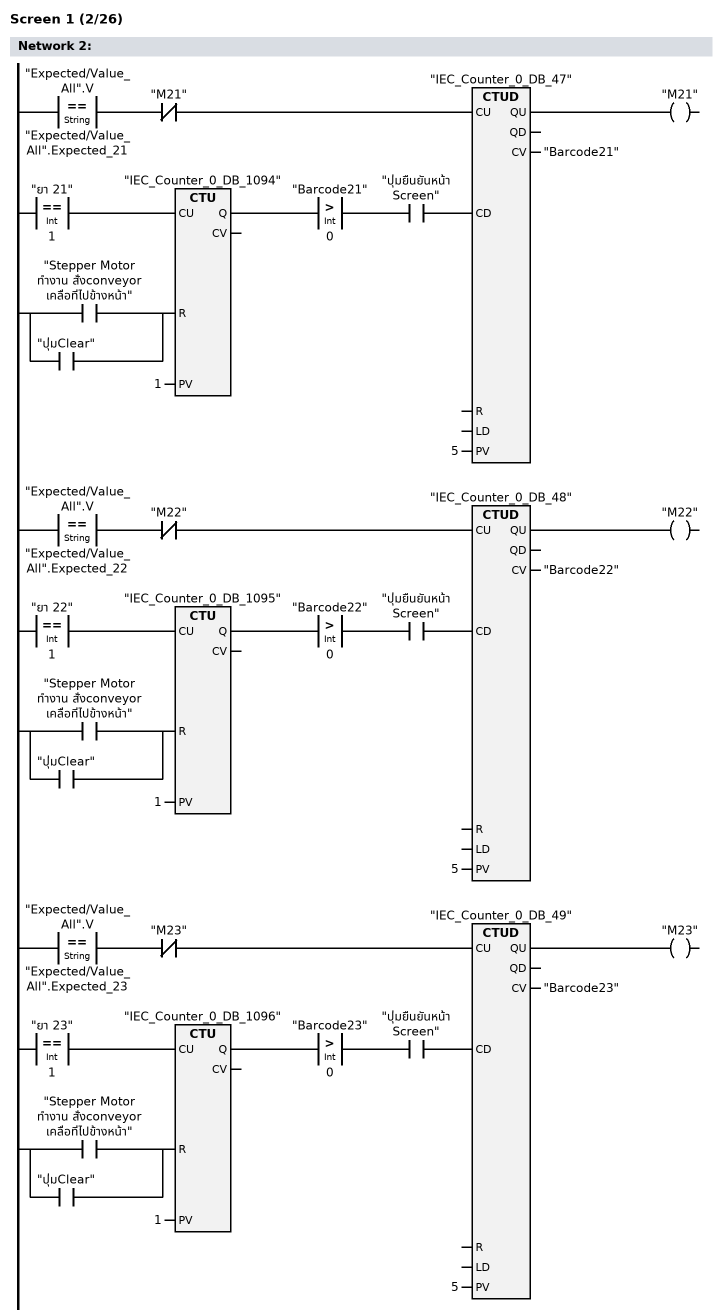
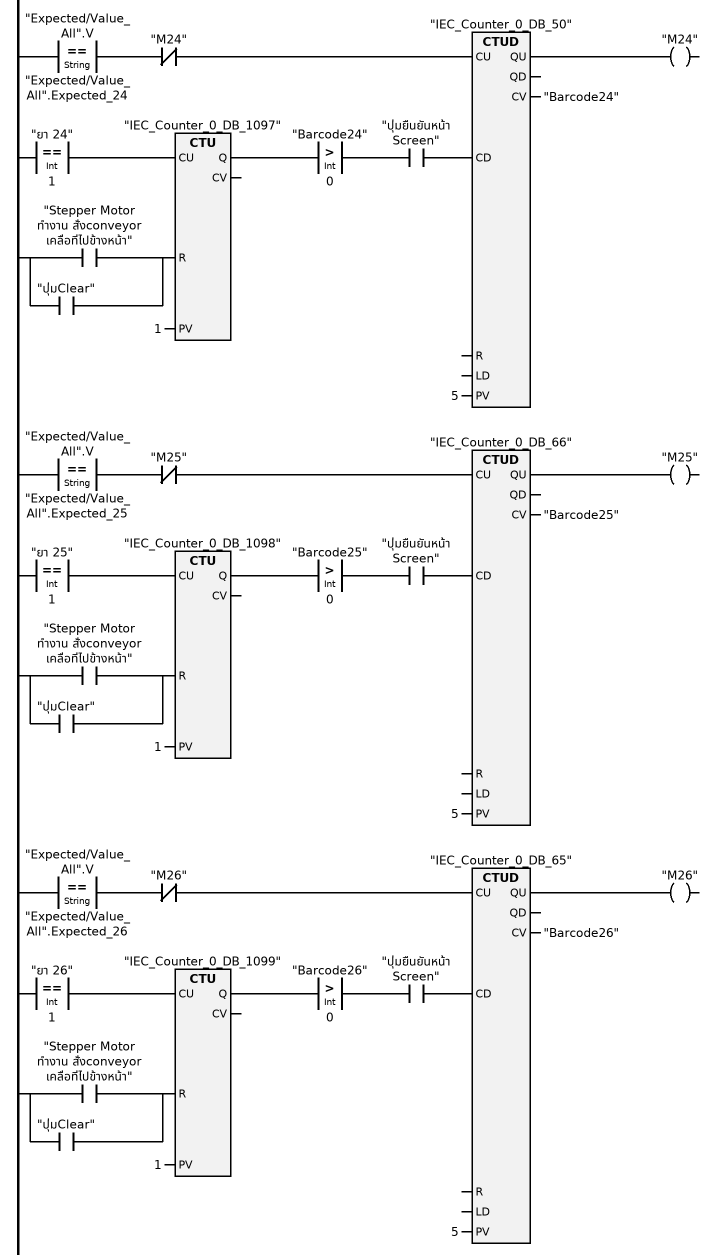
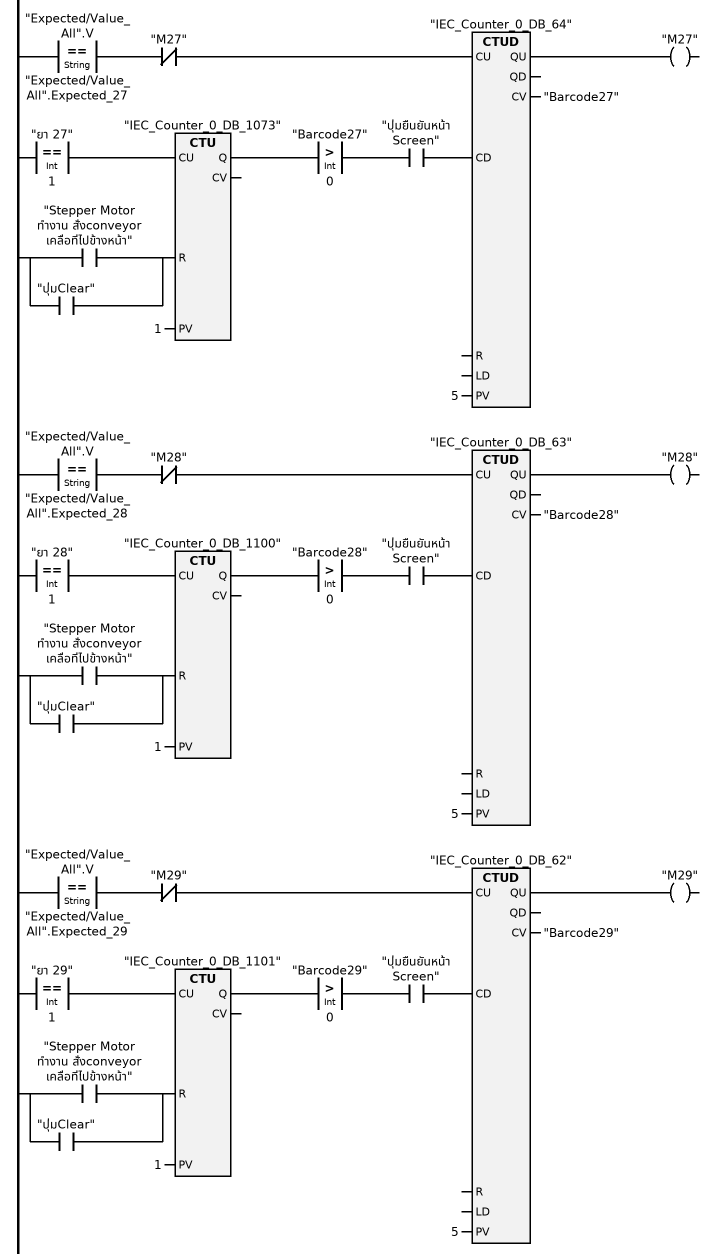
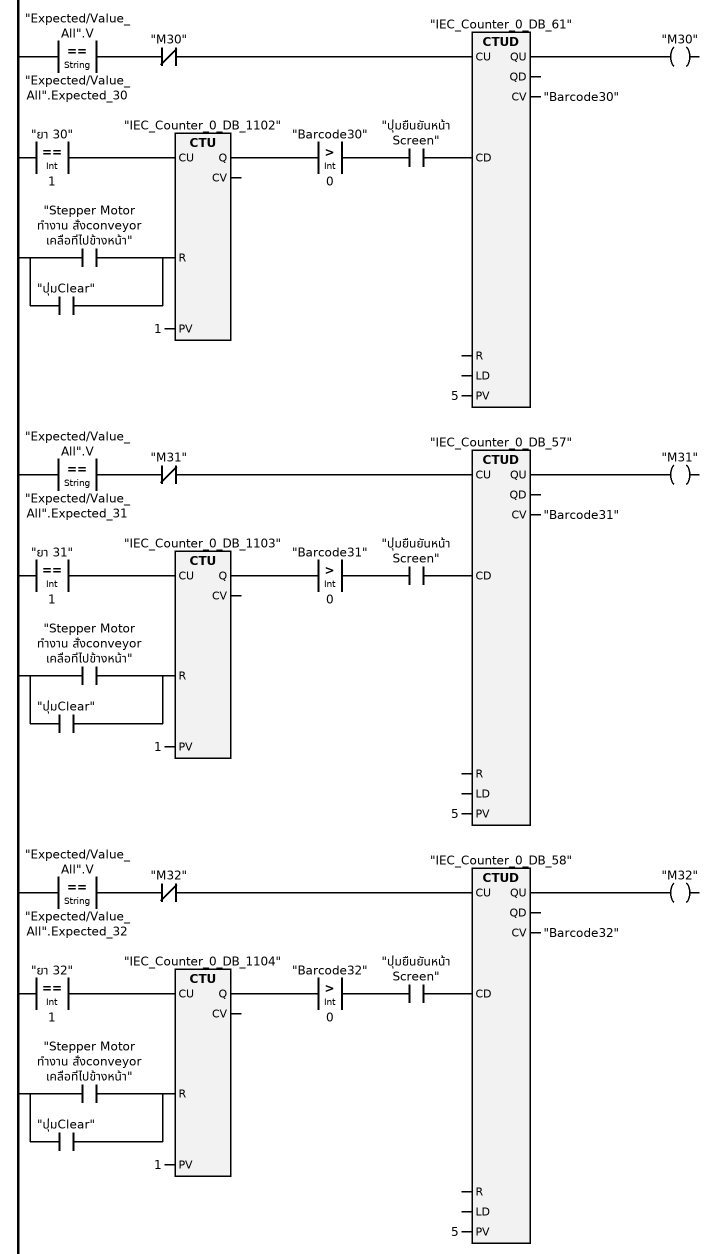
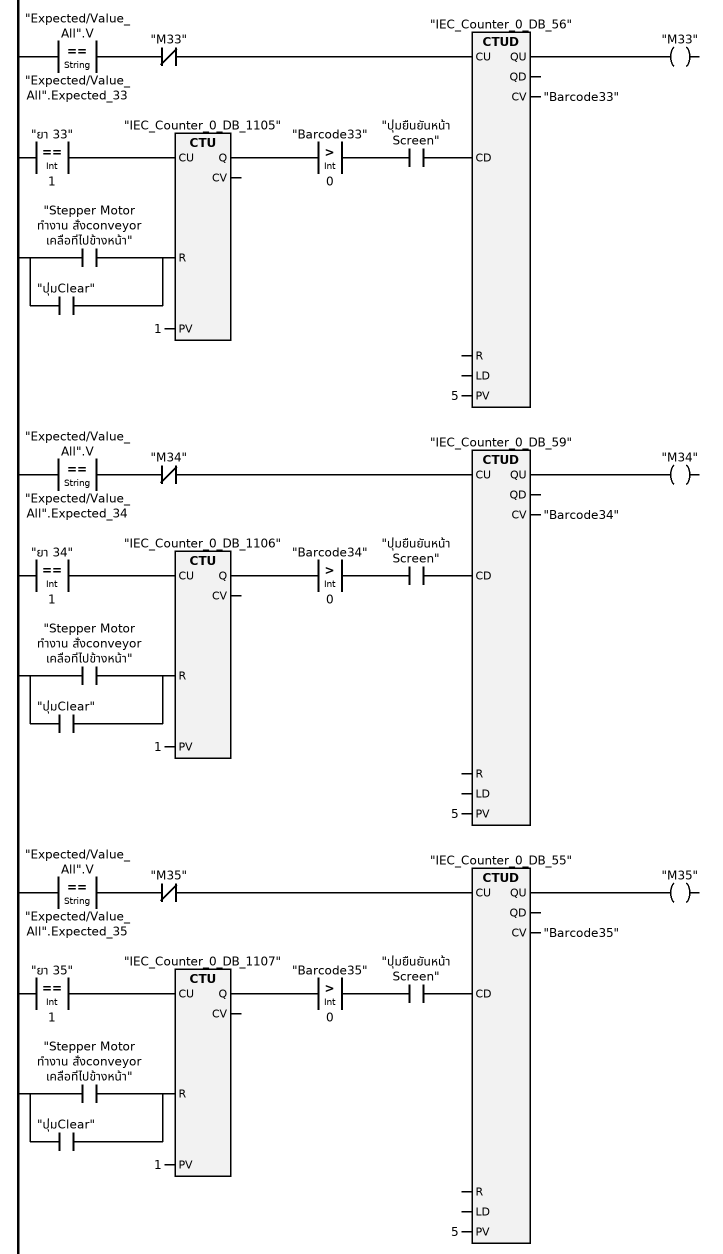
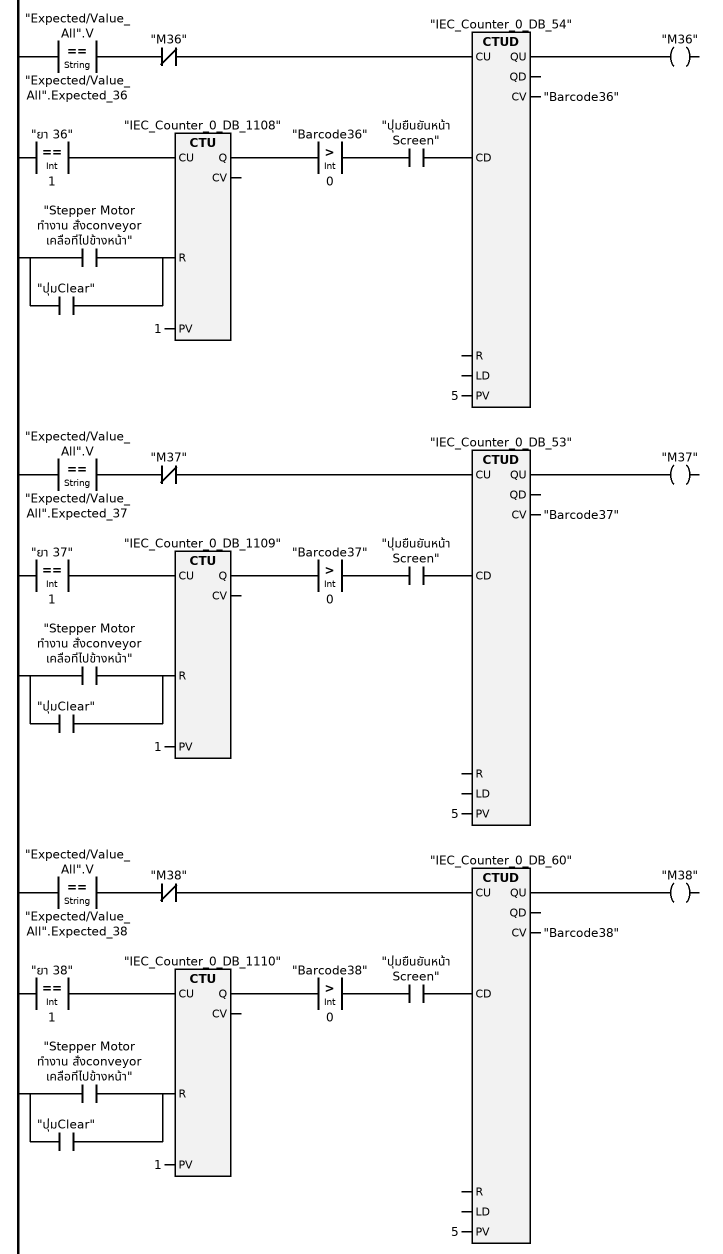
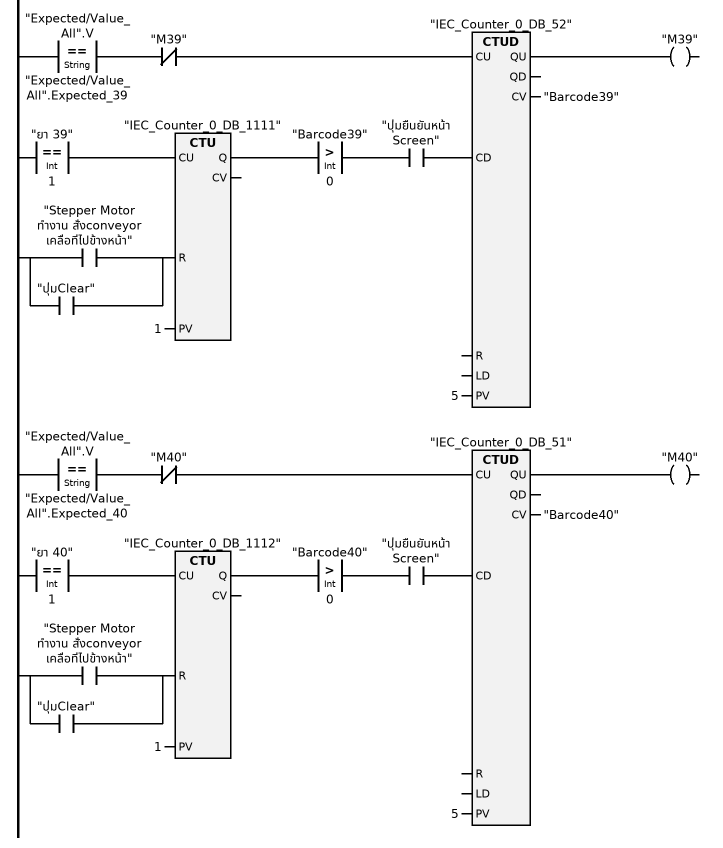
   "IEC_Counter_0_DB_1094".CTU(CU := "ยา 21" = 1,
                           R := "Stepper Motor ทำงาน สั่งconveyor เคลื่อที่ไปข้างหน้า" OR "ปุ่มClear",
                           PV := 1);
   "IEC_Counter_0_DB_47".CTUD(CU := ("Expected/Value_All".V = "Expected/Value_All".Expected_21) AND NOT "M21",
                           CD := "IEC_Counter_0_DB_1094".Q AND ("Barcode21" > 0) AND "ปุ่มยืนยันหน้า Screen",
                           PV := 5,
                           CV => "Barcode21");
   "M21" := "IEC_Counter_0_DB_47".QU;
   "IEC_Counter_0_DB_1095".CTU(CU := "ยา 22" = 1,
                           R := "Stepper Motor ทำงาน สั่งconveyor เคลื่อที่ไปข้างหน้า" OR "ปุ่มClear",
                           PV := 1);
   "IEC_Counter_0_DB_48".CTUD(CU := ("Expected/Value_All".V = "Expected/Value_All".Expected_22) AND NOT "M22",
                           CD := "IEC_Counter_0_DB_1095".Q AND ("Barcode22" > 0) AND "ปุ่มยืนยันหน้า Screen",
                           PV := 5,
                           CV => "Barcode22");
   "M22" := "IEC_Counter_0_DB_48".QU;
   "IEC_Counter_0_DB_1096".CTU(CU := "ยา 23" = 1,
                           R := "Stepper Motor ทำงาน สั่งconveyor เคลื่อที่ไปข้างหน้า" OR "ปุ่มClear",
                           PV := 1);
   "IEC_Counter_0_DB_49".CTUD(CU := ("Expected/Value_All".V = "Expected/Value_All".Expected_23) AND NOT "M23",
                           CD := "IEC_Counter_0_DB_1096".Q AND ("Barcode23" > 0) AND "ปุ่มยืนยันหน้า Screen",
                           PV := 5,
                           CV => "Barcode23");
   "M23" := "IEC_Counter_0_DB_49".QU;
   "IEC_Counter_0_DB_1097".CTU(CU := "ยา 24" = 1,
                           R := "Stepper Motor ทำงาน สั่งconveyor เคลื่อที่ไปข้างหน้า" OR "ปุ่มClear",
                           PV := 1);
   "IEC_Counter_0_DB_50".CTUD(CU := ("Expected/Value_All".V = "Expected/Value_All".Expected_24) AND NOT "M24",
                           CD := "IEC_Counter_0_DB_1097".Q AND ("Barcode24" > 0) AND "ปุ่มยืนยันหน้า Screen",
                           PV := 5,
                           CV => "Barcode24");
   "M24" := "IEC_Counter_0_DB_50".QU;
   "IEC_Counter_0_DB_1098".CTU(CU := "ยา 25" = 1,
                           R := "Stepper Motor ทำงาน สั่งconveyor เคลื่อที่ไปข้างหน้า" OR "ปุ่มClear",
                           PV := 1);
   "IEC_Counter_0_DB_66".CTUD(CU := ("Expected/Value_All".V = "Expected/Value_All".Expected_25) AND NOT "M25",
                           CD := "IEC_Counter_0_DB_1098".Q AND ("Barcode25" > 0) AND "ปุ่มยืนยันหน้า Screen",
                           PV := 5,
                           CV => "Barcode25");
   "M25" := "IEC_Counter_0_DB_66".QU;
   "IEC_Counter_0_DB_1099".CTU(CU := "ยา 26" = 1,
                           R := "Stepper Motor ทำงาน สั่งconveyor เคลื่อที่ไปข้างหน้า" OR "ปุ่มClear",
                           PV := 1);
   "IEC_Counter_0_DB_65".CTUD(CU := ("Expected/Value_All".V = "Expected/Value_All".Expected_26) AND NOT "M26",
                           CD := "IEC_Counter_0_DB_1099".Q AND ("Barcode26" > 0) AND "ปุ่มยืนยันหน้า Screen",
                           PV := 5,
                           CV => "Barcode26");
   "M26" := "IEC_Counter_0_DB_65".QU;
   "IEC_Counter_0_DB_1073".CTU(CU := "ยา 27" = 1,
                           R := "Stepper Motor ทำงาน สั่งconveyor เคลื่อที่ไปข้างหน้า" OR "ปุ่มClear",
                           PV := 1);
   "IEC_Counter_0_DB_64".CTUD(CU := ("Expected/Value_All".V = "Expected/Value_All".Expected_27) AND NOT "M27",
                           CD := "IEC_Counter_0_DB_1073".Q AND ("Barcode27" > 0) AND "ปุ่มยืนยันหน้า Screen",
                           PV := 5,
                           CV => "Barcode27");
   "M27" := "IEC_Counter_0_DB_64".QU;
   "IEC_Counter_0_DB_1100".CTU(CU := "ยา 28" = 1,
                           R := "Stepper Motor ทำงาน สั่งconveyor เคลื่อที่ไปข้างหน้า" OR "ปุ่มClear",
                           PV := 1);
   "IEC_Counter_0_DB_63".CTUD(CU := ("Expected/Value_All".V = "Expected/Value_All".Expected_28) AND NOT "M28",
                           CD := "IEC_Counter_0_DB_1100".Q AND ("Barcode28" > 0) AND "ปุ่มยืนยันหน้า Screen",
                           PV := 5,
                           CV => "Barcode28");
   "M28" := "IEC_Counter_0_DB_63".QU;
   "IEC_Counter_0_DB_1101".CTU(CU := "ยา 29" = 1,
                           R := "Stepper Motor ทำงาน สั่งconveyor เคลื่อที่ไปข้างหน้า" OR "ปุ่มClear",
                           PV := 1);
   "IEC_Counter_0_DB_62".CTUD(CU := ("Expected/Value_All".V = "Expected/Value_All".Expected_29) AND NOT "M29",
                           CD := "IEC_Counter_0_DB_1101".Q AND ("Barcode29" > 0) AND "ปุ่มยืนยันหน้า Screen",
                           PV := 5,
                           CV => "Barcode29");
   "M29" := "IEC_Counter_0_DB_62".QU;
   "IEC_Counter_0_DB_1102".CTU(CU := "ยา 30" = 1,
                           R := "Stepper Motor ทำงาน สั่งconveyor เคลื่อที่ไปข้างหน้า" OR "ปุ่มClear",
                           PV := 1);
   "IEC_Counter_0_DB_61".CTUD(CU := ("Expected/Value_All".V = "Expected/Value_All".Expected_30) AND NOT "M30",
                           CD := "IEC_Counter_0_DB_1102".Q AND ("Barcode30" > 0) AND "ปุ่มยืนยันหน้า Screen",
                           PV := 5,
                           CV => "Barcode30");
   "M30" := "IEC_Counter_0_DB_61".QU;
   "IEC_Counter_0_DB_1103".CTU(CU := "ยา 31" = 1,
                           R := "Stepper Motor ทำงาน สั่งconveyor เคลื่อที่ไปข้างหน้า" OR "ปุ่มClear",
                           PV := 1);
   "IEC_Counter_0_DB_57".CTUD(CU := ("Expected/Value_All".V = "Expected/Value_All".Expected_31) AND NOT "M31",
                           CD := "IEC_Counter_0_DB_1103".Q AND ("Barcode31" > 0) AND "ปุ่มยืนยันหน้า Screen",
                           PV := 5,
                           CV => "Barcode31");
   "M31" := "IEC_Counter_0_DB_57".QU;
   "IEC_Counter_0_DB_1104".CTU(CU := "ยา 32" = 1,
                           R := "Stepper Motor ทำงาน สั่งconveyor เคลื่อที่ไปข้างหน้า" OR "ปุ่มClear",
                           PV := 1);
   "IEC_Counter_0_DB_58".CTUD(CU := ("Expected/Value_All".V = "Expected/Value_All".Expected_32) AND NOT "M32",
                           CD := "IEC_Counter_0_DB_1104".Q AND ("Barcode32" > 0) AND "ปุ่มยืนยันหน้า Screen",
                           PV := 5,
                           CV => "Barcode32");
   "M32" := "IEC_Counter_0_DB_58".QU;
   "IEC_Counter_0_DB_1105".CTU(CU := "ยา 33" = 1,
                           R := "Stepper Motor ทำงาน สั่งconveyor เคลื่อที่ไปข้างหน้า" OR "ปุ่มClear",
                           PV := 1);
   "IEC_Counter_0_DB_56".CTUD(CU := ("Expected/Value_All".V = "Expected/Value_All".Expected_33) AND NOT "M33",
                           CD := "IEC_Counter_0_DB_1105".Q AND ("Barcode33" > 0) AND "ปุ่มยืนยันหน้า Screen",
                           PV := 5,
                           CV => "Barcode33");
   "M33" := "IEC_Counter_0_DB_56".QU;
   "IEC_Counter_0_DB_1106".CTU(CU := "ยา 34" = 1,
                           R := "Stepper Motor ทำงาน สั่งconveyor เคลื่อที่ไปข้างหน้า" OR "ปุ่มClear",
                           PV := 1);
   "IEC_Counter_0_DB_59".CTUD(CU := ("Expected/Value_All".V = "Expected/Value_All".Expected_34) AND NOT "M34",
                           CD := "IEC_Counter_0_DB_1106".Q AND ("Barcode34" > 0) AND "ปุ่มยืนยันหน้า Screen",
                           PV := 5,
                           CV => "Barcode34");
   "M34" := "IEC_Counter_0_DB_59".QU;
   "IEC_Counter_0_DB_1107".CTU(CU := "ยา 35" = 1,
                           R := "Stepper Motor ทำงาน สั่งconveyor เคลื่อที่ไปข้างหน้า" OR "ปุ่มClear",
                           PV := 1);
   "IEC_Counter_0_DB_55".CTUD(CU := ("Expected/Value_All".V = "Expected/Value_All".Expected_35) AND NOT "M35",
                           CD := "IEC_Counter_0_DB_1107".Q AND ("Barcode35" > 0) AND "ปุ่มยืนยันหน้า Screen",
                           PV := 5,
                           CV => "Barcode35");
   "M35" := "IEC_Counter_0_DB_55".QU;
   "IEC_Counter_0_DB_1108".CTU(CU := "ยา 36" = 1,
                           R := "Stepper Motor ทำงาน สั่งconveyor เคลื่อที่ไปข้างหน้า" OR "ปุ่มClear",
                           PV := 1);
   "IEC_Counter_0_DB_54".CTUD(CU := ("Expected/Value_All".V = "Expected/Value_All".Expected_36) AND NOT "M36",
                           CD := "IEC_Counter_0_DB_1108".Q AND ("Barcode36" > 0) AND "ปุ่มยืนยันหน้า Screen",
                           PV := 5,
                           CV => "Barcode36");
   "M36" := "IEC_Counter_0_DB_54".QU;
   "IEC_Counter_0_DB_1109".CTU(CU := "ยา 37" = 1,
                           R := "Stepper Motor ทำงาน สั่งconveyor เคลื่อที่ไปข้างหน้า" OR "ปุ่มClear",
                           PV := 1);
   "IEC_Counter_0_DB_53".CTUD(CU := ("Expected/Value_All".V = "Expected/Value_All".Expected_37) AND NOT "M37",
                           CD := "IEC_Counter_0_DB_1109".Q AND ("Barcode37" > 0) AND "ปุ่มยืนยันหน้า Screen",
                           PV := 5,
                           CV => "Barcode37");
   "M37" := "IEC_Counter_0_DB_53".QU;
   "IEC_Counter_0_DB_1110".CTU(CU := "ยา 38" = 1,
                           R := "Stepper Motor ทำงาน สั่งconveyor เคลื่อที่ไปข้างหน้า" OR "ปุ่มClear",
                           PV := 1);
   "IEC_Counter_0_DB_60".CTUD(CU := ("Expected/Value_All".V = "Expected/Value_All".Expected_38) AND NOT "M38",
                           CD := "IEC_Counter_0_DB_1110".Q AND ("Barcode38" > 0) AND "ปุ่มยืนยันหน้า Screen",
                           PV := 5,
                           CV => "Barcode38");
   "M38" := "IEC_Counter_0_DB_60".QU;
   "IEC_Counter_0_DB_1111".CTU(CU := "ยา 39" = 1,
                           R := "Stepper Motor ทำงาน สั่งconveyor เคลื่อที่ไปข้างหน้า" OR "ปุ่มClear",
                           PV := 1);
   "IEC_Counter_0_DB_52".CTUD(CU := ("Expected/Value_All".V = "Expected/Value_All".Expected_39) AND NOT "M39",
                           CD := "IEC_Counter_0_DB_1111".Q AND ("Barcode39" > 0) AND "ปุ่มยืนยันหน้า Screen",
                           PV := 5,
                           CV => "Barcode39");
   "M39" := "IEC_Counter_0_DB_52".QU;
   "IEC_Counter_0_DB_1112".CTU(CU := "ยา 40" = 1,
                           R := "Stepper Motor ทำงาน สั่งconveyor เคลื่อที่ไปข้างหน้า" OR "ปุ่มClear",
                           PV := 1);
   "IEC_Counter_0_DB_51".CTUD(CU := ("Expected/Value_All".V = "Expected/Value_All".Expected_40) AND NOT "M40",
                           CD := "IEC_Counter_0_DB_1112".Q AND ("Barcode40" > 0) AND "ปุ่มยืนยันหน้า Screen",
                           PV := 5,
                           CV => "Barcode40");
   "M40" := "IEC_Counter_0_DB_51".QU;
END_REGION

REGION Network 3
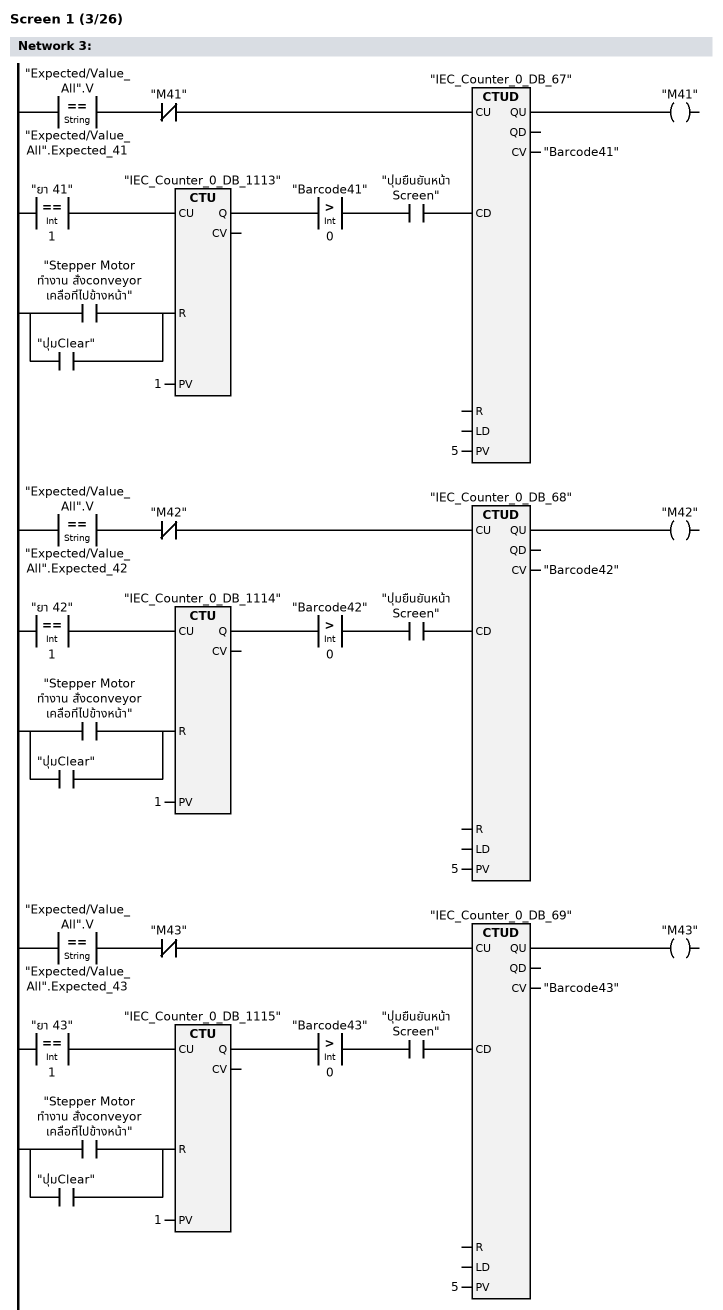
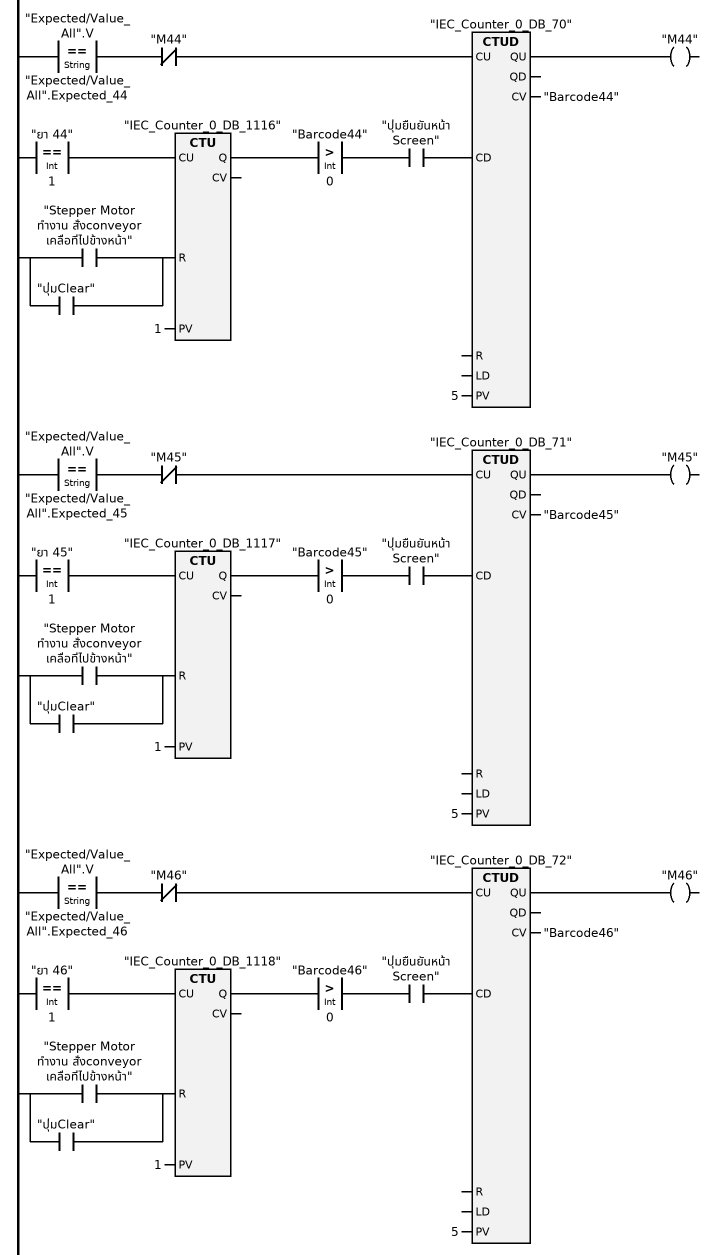
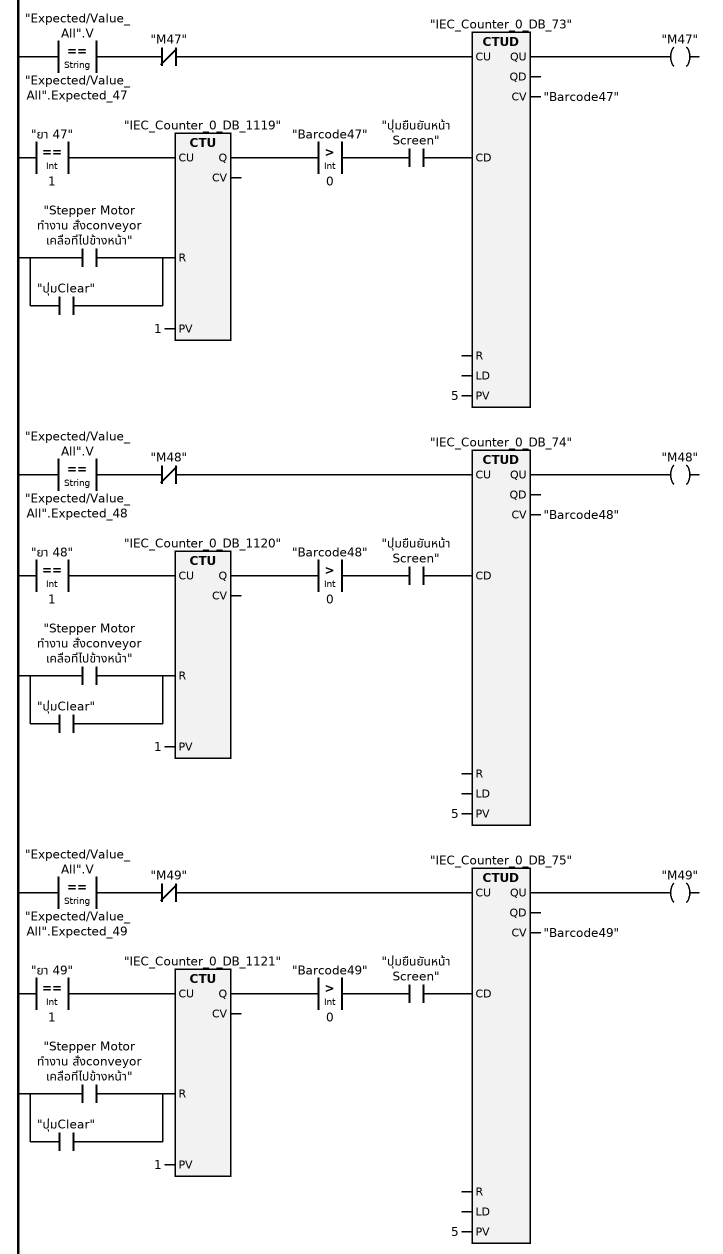
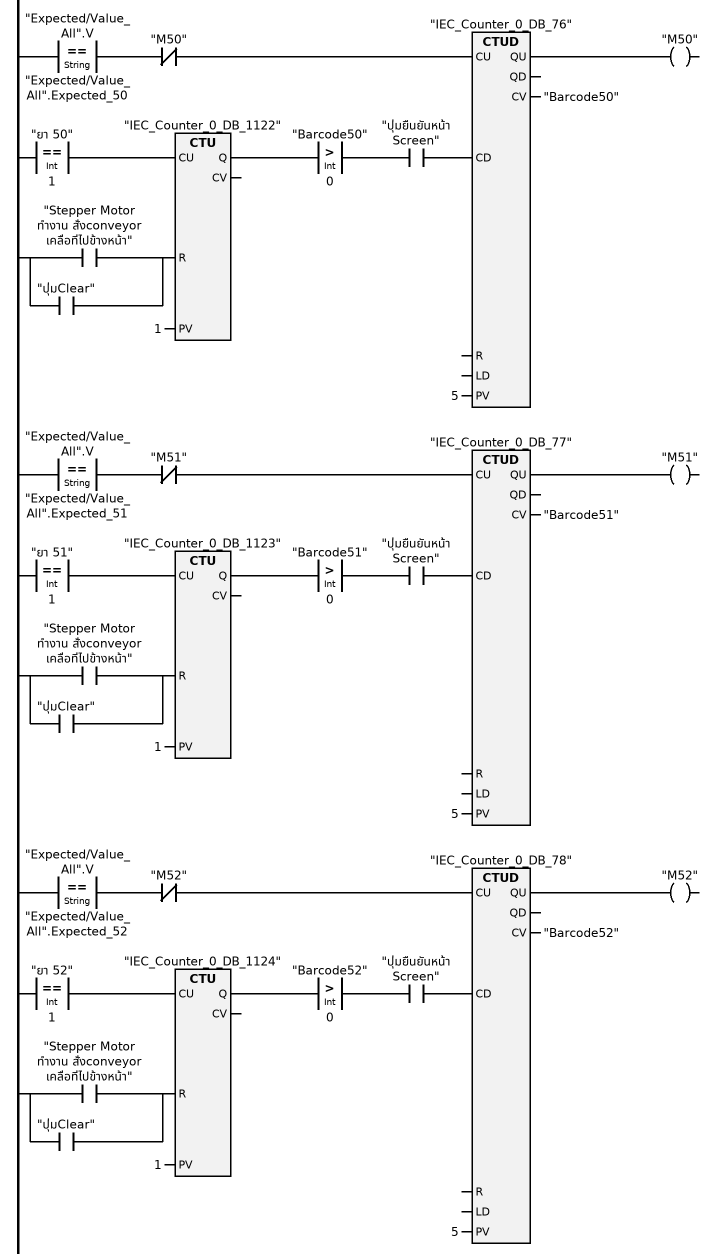
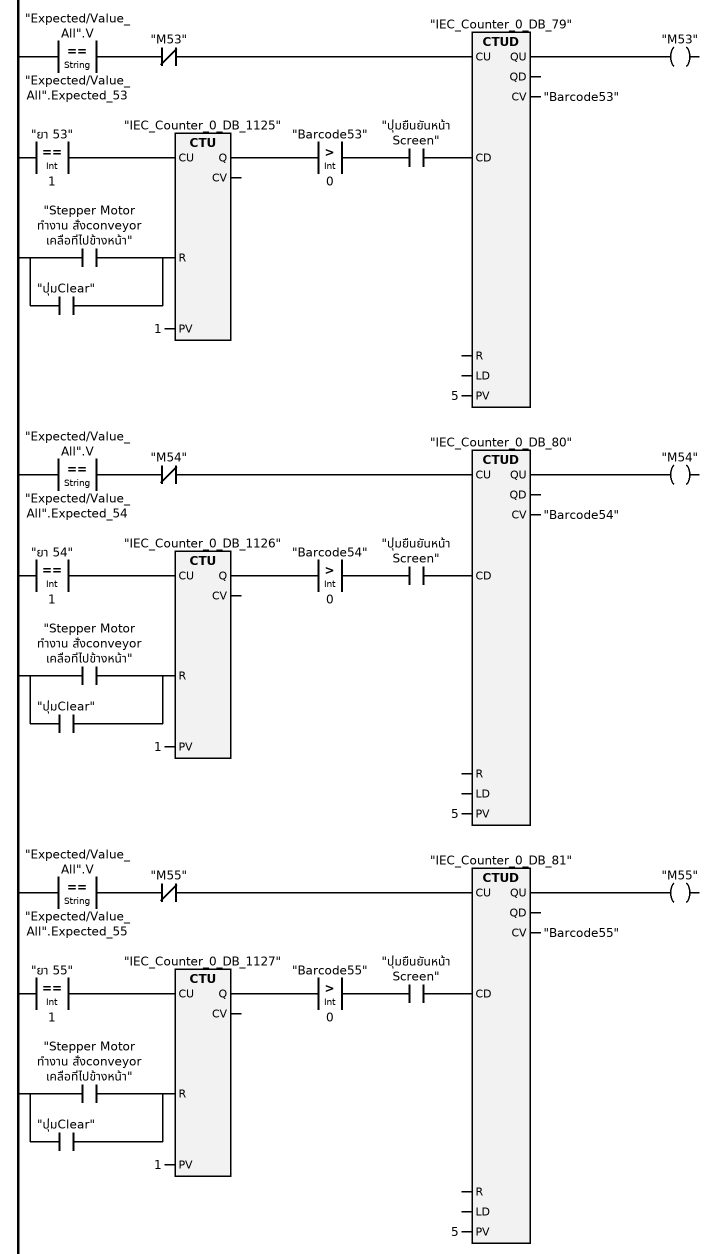
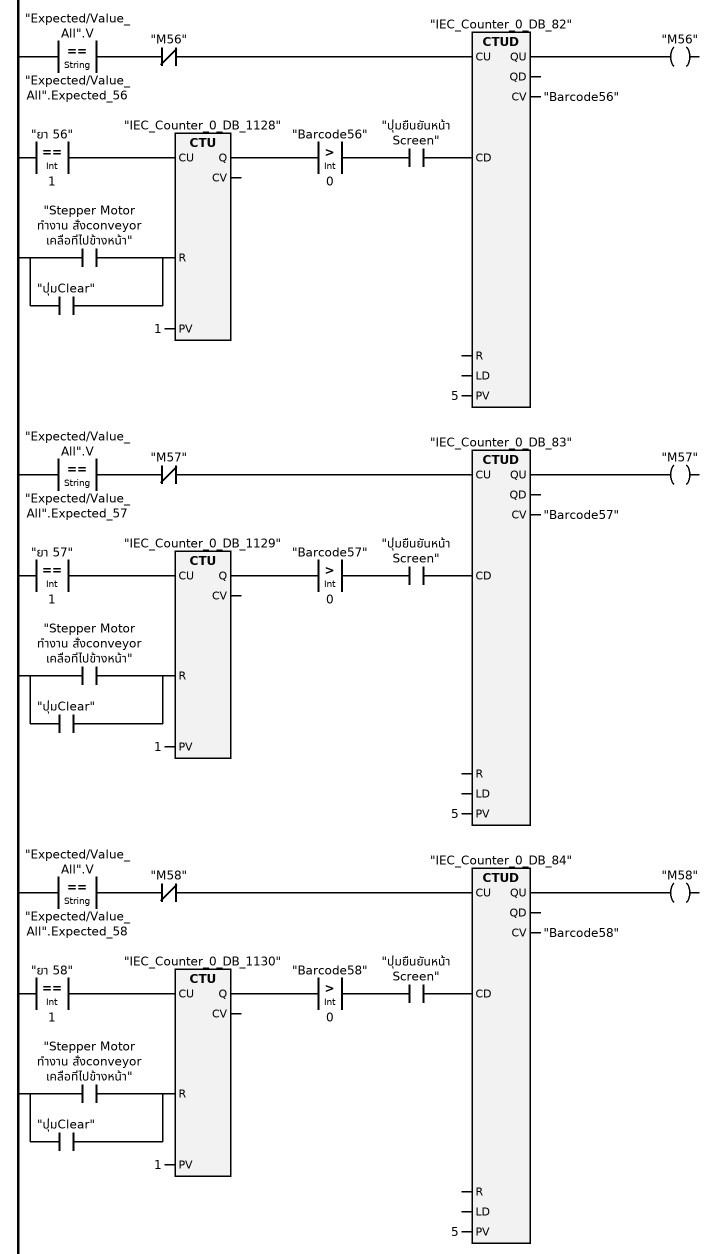
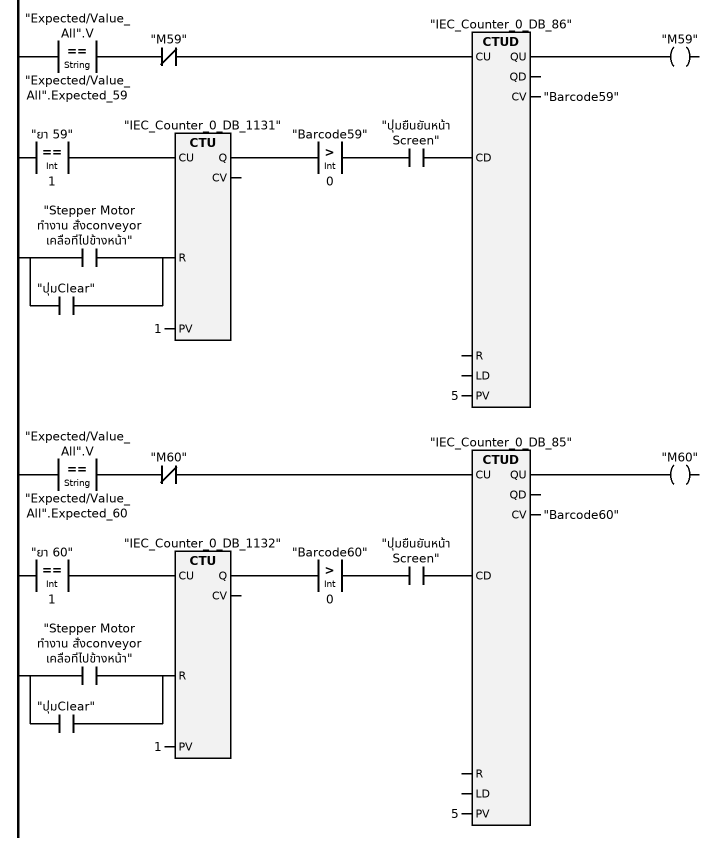
   "IEC_Counter_0_DB_1113".CTU(CU := "ยา 41" = 1,
                           R := "Stepper Motor ทำงาน สั่งconveyor เคลื่อที่ไปข้างหน้า" OR "ปุ่มClear",
                           PV := 1);
   "IEC_Counter_0_DB_67".CTUD(CU := ("Expected/Value_All".V = "Expected/Value_All".Expected_41) AND NOT "M41",
                           CD := "IEC_Counter_0_DB_1113".Q AND ("Barcode41" > 0) AND "ปุ่มยืนยันหน้า Screen",
                           PV := 5,
                           CV => "Barcode41");
   "M41" := "IEC_Counter_0_DB_67".QU;
   "IEC_Counter_0_DB_1114".CTU(CU := "ยา 42" = 1,
                           R := "Stepper Motor ทำงาน สั่งconveyor เคลื่อที่ไปข้างหน้า" OR "ปุ่มClear",
                           PV := 1);
   "IEC_Counter_0_DB_68".CTUD(CU := ("Expected/Value_All".V = "Expected/Value_All".Expected_42) AND NOT "M42",
                           CD := "IEC_Counter_0_DB_1114".Q AND ("Barcode42" > 0) AND "ปุ่มยืนยันหน้า Screen",
                           PV := 5,
                           CV => "Barcode42");
   "M42" := "IEC_Counter_0_DB_68".QU;
   "IEC_Counter_0_DB_1115".CTU(CU := "ยา 43" = 1,
                           R := "Stepper Motor ทำงาน สั่งconveyor เคลื่อที่ไปข้างหน้า" OR "ปุ่มClear",
                           PV := 1);
   "IEC_Counter_0_DB_69".CTUD(CU := ("Expected/Value_All".V = "Expected/Value_All".Expected_43) AND NOT "M43",
                           CD := "IEC_Counter_0_DB_1115".Q AND ("Barcode43" > 0) AND "ปุ่มยืนยันหน้า Screen",
                           PV := 5,
                           CV => "Barcode43");
   "M43" := "IEC_Counter_0_DB_69".QU;
   "IEC_Counter_0_DB_1116".CTU(CU := "ยา 44" = 1,
                           R := "Stepper Motor ทำงาน สั่งconveyor เคลื่อที่ไปข้างหน้า" OR "ปุ่มClear",
                           PV := 1);
   "IEC_Counter_0_DB_70".CTUD(CU := ("Expected/Value_All".V = "Expected/Value_All".Expected_44) AND NOT "M44",
                           CD := "IEC_Counter_0_DB_1116".Q AND ("Barcode44" > 0) AND "ปุ่มยืนยันหน้า Screen",
                           PV := 5,
                           CV => "Barcode44");
   "M44" := "IEC_Counter_0_DB_70".QU;
   "IEC_Counter_0_DB_1117".CTU(CU := "ยา 45" = 1,
                           R := "Stepper Motor ทำงาน สั่งconveyor เคลื่อที่ไปข้างหน้า" OR "ปุ่มClear",
                           PV := 1);
   "IEC_Counter_0_DB_71".CTUD(CU := ("Expected/Value_All".V = "Expected/Value_All".Expected_45) AND NOT "M45",
                           CD := "IEC_Counter_0_DB_1117".Q AND ("Barcode45" > 0) AND "ปุ่มยืนยันหน้า Screen",
                           PV := 5,
                           CV => "Barcode45");
   "M45" := "IEC_Counter_0_DB_71".QU;
   "IEC_Counter_0_DB_1118".CTU(CU := "ยา 46" = 1,
                           R := "Stepper Motor ทำงาน สั่งconveyor เคลื่อที่ไปข้างหน้า" OR "ปุ่มClear",
                           PV := 1);
   "IEC_Counter_0_DB_72".CTUD(CU := ("Expected/Value_All".V = "Expected/Value_All".Expected_46) AND NOT "M46",
                           CD := "IEC_Counter_0_DB_1118".Q AND ("Barcode46" > 0) AND "ปุ่มยืนยันหน้า Screen",
                           PV := 5,
                           CV => "Barcode46");
   "M46" := "IEC_Counter_0_DB_72".QU;
   "IEC_Counter_0_DB_1119".CTU(CU := "ยา 47" = 1,
                           R := "Stepper Motor ทำงาน สั่งconveyor เคลื่อที่ไปข้างหน้า" OR "ปุ่มClear",
                           PV := 1);
   "IEC_Counter_0_DB_73".CTUD(CU := ("Expected/Value_All".V = "Expected/Value_All".Expected_47) AND NOT "M47",
                           CD := "IEC_Counter_0_DB_1119".Q AND ("Barcode47" > 0) AND "ปุ่มยืนยันหน้า Screen",
                           PV := 5,
                           CV => "Barcode47");
   "M47" := "IEC_Counter_0_DB_73".QU;
   "IEC_Counter_0_DB_1120".CTU(CU := "ยา 48" = 1,
                           R := "Stepper Motor ทำงาน สั่งconveyor เคลื่อที่ไปข้างหน้า" OR "ปุ่มClear",
                           PV := 1);
   "IEC_Counter_0_DB_74".CTUD(CU := ("Expected/Value_All".V = "Expected/Value_All".Expected_48) AND NOT "M48",
                           CD := "IEC_Counter_0_DB_1120".Q AND ("Barcode48" > 0) AND "ปุ่มยืนยันหน้า Screen",
                           PV := 5,
                           CV => "Barcode48");
   "M48" := "IEC_Counter_0_DB_74".QU;
   "IEC_Counter_0_DB_1121".CTU(CU := "ยา 49" = 1,
                           R := "Stepper Motor ทำงาน สั่งconveyor เคลื่อที่ไปข้างหน้า" OR "ปุ่มClear",
                           PV := 1);
   "IEC_Counter_0_DB_75".CTUD(CU := ("Expected/Value_All".V = "Expected/Value_All".Expected_49) AND NOT "M49",
                           CD := "IEC_Counter_0_DB_1121".Q AND ("Barcode49" > 0) AND "ปุ่มยืนยันหน้า Screen",
                           PV := 5,
                           CV => "Barcode49");
   "M49" := "IEC_Counter_0_DB_75".QU;
   "IEC_Counter_0_DB_1122".CTU(CU := "ยา 50" = 1,
                           R := "Stepper Motor ทำงาน สั่งconveyor เคลื่อที่ไปข้างหน้า" OR "ปุ่มClear",
                           PV := 1);
   "IEC_Counter_0_DB_76".CTUD(CU := ("Expected/Value_All".V = "Expected/Value_All".Expected_50) AND NOT "M50",
                           CD := "IEC_Counter_0_DB_1122".Q AND ("Barcode50" > 0) AND "ปุ่มยืนยันหน้า Screen",
                           PV := 5,
                           CV => "Barcode50");
   "M50" := "IEC_Counter_0_DB_76".QU;
   "IEC_Counter_0_DB_1123".CTU(CU := "ยา 51" = 1,
                           R := "Stepper Motor ทำงาน สั่งconveyor เคลื่อที่ไปข้างหน้า" OR "ปุ่มClear",
                           PV := 1);
   "IEC_Counter_0_DB_77".CTUD(CU := ("Expected/Value_All".V = "Expected/Value_All".Expected_51) AND NOT "M51",
                           CD := "IEC_Counter_0_DB_1123".Q AND ("Barcode51" > 0) AND "ปุ่มยืนยันหน้า Screen",
                           PV := 5,
                           CV => "Barcode51");
   "M51" := "IEC_Counter_0_DB_77".QU;
   "IEC_Counter_0_DB_1124".CTU(CU := "ยา 52" = 1,
                           R := "Stepper Motor ทำงาน สั่งconveyor เคลื่อที่ไปข้างหน้า" OR "ปุ่มClear",
                           PV := 1);
   "IEC_Counter_0_DB_78".CTUD(CU := ("Expected/Value_All".V = "Expected/Value_All".Expected_52) AND NOT "M52",
                           CD := "IEC_Counter_0_DB_1124".Q AND ("Barcode52" > 0) AND "ปุ่มยืนยันหน้า Screen",
                           PV := 5,
                           CV => "Barcode52");
   "M52" := "IEC_Counter_0_DB_78".QU;
   "IEC_Counter_0_DB_1125".CTU(CU := "ยา 53" = 1,
                           R := "Stepper Motor ทำงาน สั่งconveyor เคลื่อที่ไปข้างหน้า" OR "ปุ่มClear",
                           PV := 1);
   "IEC_Counter_0_DB_79".CTUD(CU := ("Expected/Value_All".V = "Expected/Value_All".Expected_53) AND NOT "M53",
                           CD := "IEC_Counter_0_DB_1125".Q AND ("Barcode53" > 0) AND "ปุ่มยืนยันหน้า Screen",
                           PV := 5,
                           CV => "Barcode53");
   "M53" := "IEC_Counter_0_DB_79".QU;
   "IEC_Counter_0_DB_1126".CTU(CU := "ยา 54" = 1,
                           R := "Stepper Motor ทำงาน สั่งconveyor เคลื่อที่ไปข้างหน้า" OR "ปุ่มClear",
                           PV := 1);
   "IEC_Counter_0_DB_80".CTUD(CU := ("Expected/Value_All".V = "Expected/Value_All".Expected_54) AND NOT "M54",
                           CD := "IEC_Counter_0_DB_1126".Q AND ("Barcode54" > 0) AND "ปุ่มยืนยันหน้า Screen",
                           PV := 5,
                           CV => "Barcode54");
   "M54" := "IEC_Counter_0_DB_80".QU;
   "IEC_Counter_0_DB_1127".CTU(CU := "ยา 55" = 1,
                           R := "Stepper Motor ทำงาน สั่งconveyor เคลื่อที่ไปข้างหน้า" OR "ปุ่มClear",
                           PV := 1);
   "IEC_Counter_0_DB_81".CTUD(CU := ("Expected/Value_All".V = "Expected/Value_All".Expected_55) AND NOT "M55",
                           CD := "IEC_Counter_0_DB_1127".Q AND ("Barcode55" > 0) AND "ปุ่มยืนยันหน้า Screen",
                           PV := 5,
                           CV => "Barcode55");
   "M55" := "IEC_Counter_0_DB_81".QU;
   "IEC_Counter_0_DB_1128".CTU(CU := "ยา 56" = 1,
                           R := "Stepper Motor ทำงาน สั่งconveyor เคลื่อที่ไปข้างหน้า" OR "ปุ่มClear",
                           PV := 1);
   "IEC_Counter_0_DB_82".CTUD(CU := ("Expected/Value_All".V = "Expected/Value_All".Expected_56) AND NOT "M56",
                           CD := "IEC_Counter_0_DB_1128".Q AND ("Barcode56" > 0) AND "ปุ่มยืนยันหน้า Screen",
                           PV := 5,
                           CV => "Barcode56");
   "M56" := "IEC_Counter_0_DB_82".QU;
   "IEC_Counter_0_DB_1129".CTU(CU := "ยา 57" = 1,
                           R := "Stepper Motor ทำงาน สั่งconveyor เคลื่อที่ไปข้างหน้า" OR "ปุ่มClear",
                           PV := 1);
   "IEC_Counter_0_DB_83".CTUD(CU := ("Expected/Value_All".V = "Expected/Value_All".Expected_57) AND NOT "M57",
                           CD := "IEC_Counter_0_DB_1129".Q AND ("Barcode57" > 0) AND "ปุ่มยืนยันหน้า Screen",
                           PV := 5,
                           CV => "Barcode57");
   "M57" := "IEC_Counter_0_DB_83".QU;
   "IEC_Counter_0_DB_1130".CTU(CU := "ยา 58" = 1,
                           R := "Stepper Motor ทำงาน สั่งconveyor เคลื่อที่ไปข้างหน้า" OR "ปุ่มClear",
                           PV := 1);
   "IEC_Counter_0_DB_84".CTUD(CU := ("Expected/Value_All".V = "Expected/Value_All".Expected_58) AND NOT "M58",
                           CD := "IEC_Counter_0_DB_1130".Q AND ("Barcode58" > 0) AND "ปุ่มยืนยันหน้า Screen",
                           PV := 5,
                           CV => "Barcode58");
   "M58" := "IEC_Counter_0_DB_84".QU;
   "IEC_Counter_0_DB_1131".CTU(CU := "ยา 59" = 1,
                           R := "Stepper Motor ทำงาน สั่งconveyor เคลื่อที่ไปข้างหน้า" OR "ปุ่มClear",
                           PV := 1);
   "IEC_Counter_0_DB_86".CTUD(CU := ("Expected/Value_All".V = "Expected/Value_All".Expected_59) AND NOT "M59",
                           CD := "IEC_Counter_0_DB_1131".Q AND ("Barcode59" > 0) AND "ปุ่มยืนยันหน้า Screen",
                           PV := 5,
                           CV => "Barcode59");
   "M59" := "IEC_Counter_0_DB_86".QU;
   "IEC_Counter_0_DB_1132".CTU(CU := "ยา 60" = 1,
                           R := "Stepper Motor ทำงาน สั่งconveyor เคลื่อที่ไปข้างหน้า" OR "ปุ่มClear",
                           PV := 1);
   "IEC_Counter_0_DB_85".CTUD(CU := ("Expected/Value_All".V = "Expected/Value_All".Expected_60) AND NOT "M60",
                           CD := "IEC_Counter_0_DB_1132".Q AND ("Barcode60" > 0) AND "ปุ่มยืนยันหน้า Screen",
                           PV := 5,
                           CV => "Barcode60");
   "M60" := "IEC_Counter_0_DB_85".QU;
END_REGION

REGION Network 4
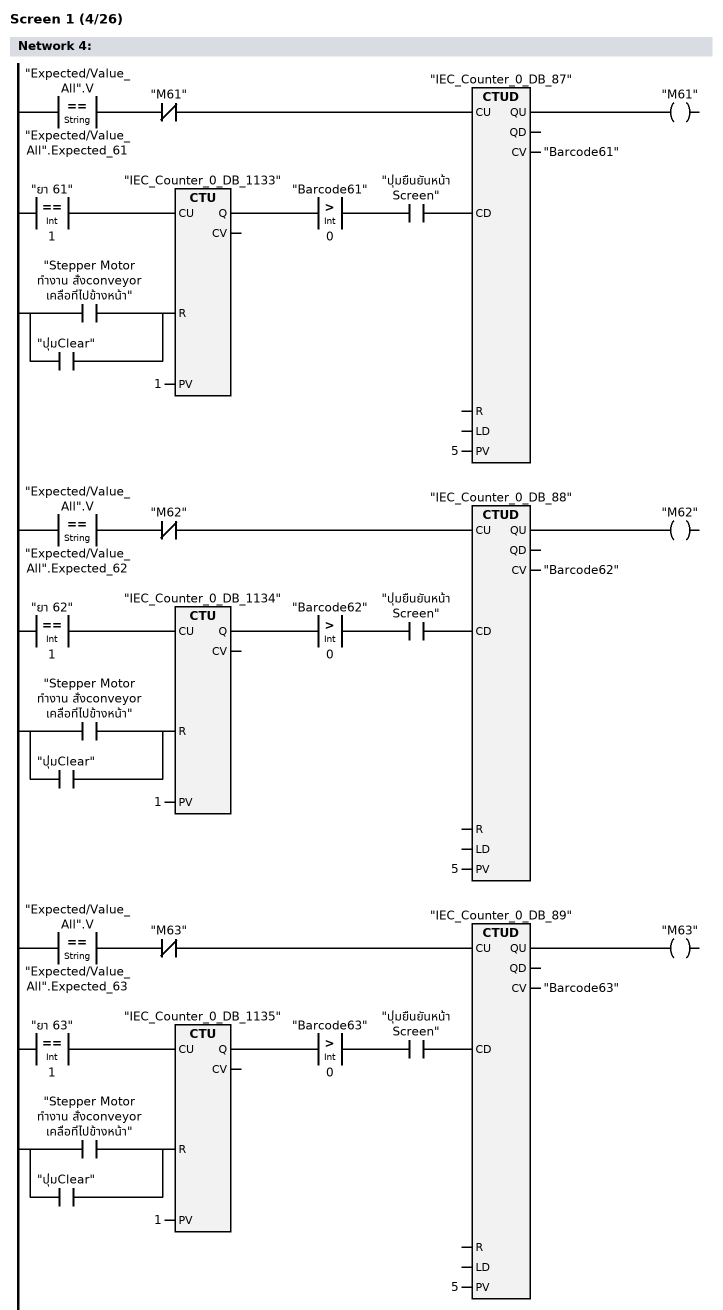
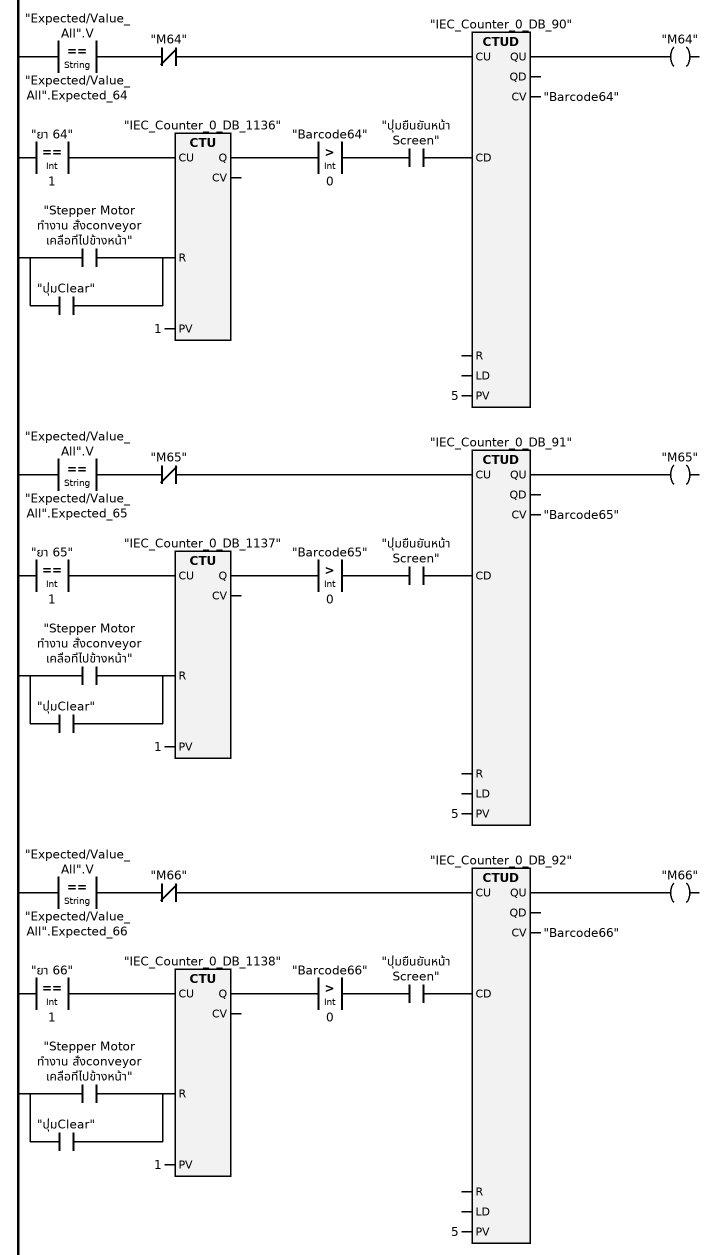
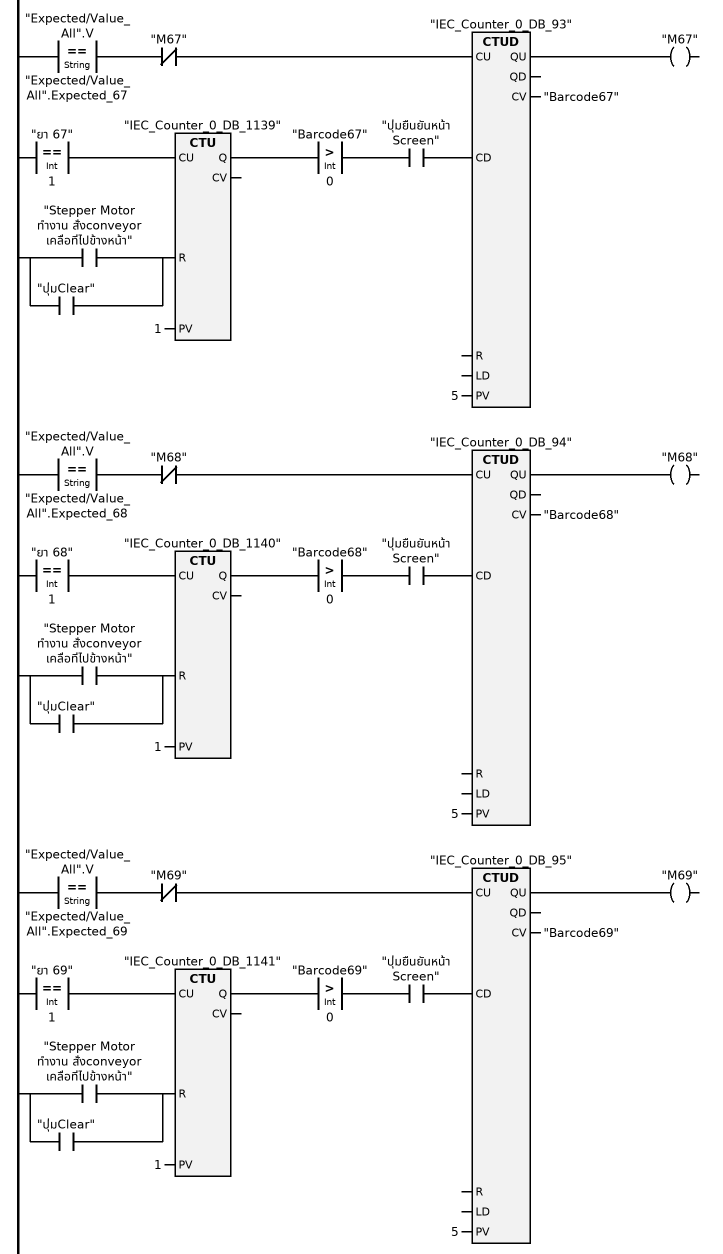
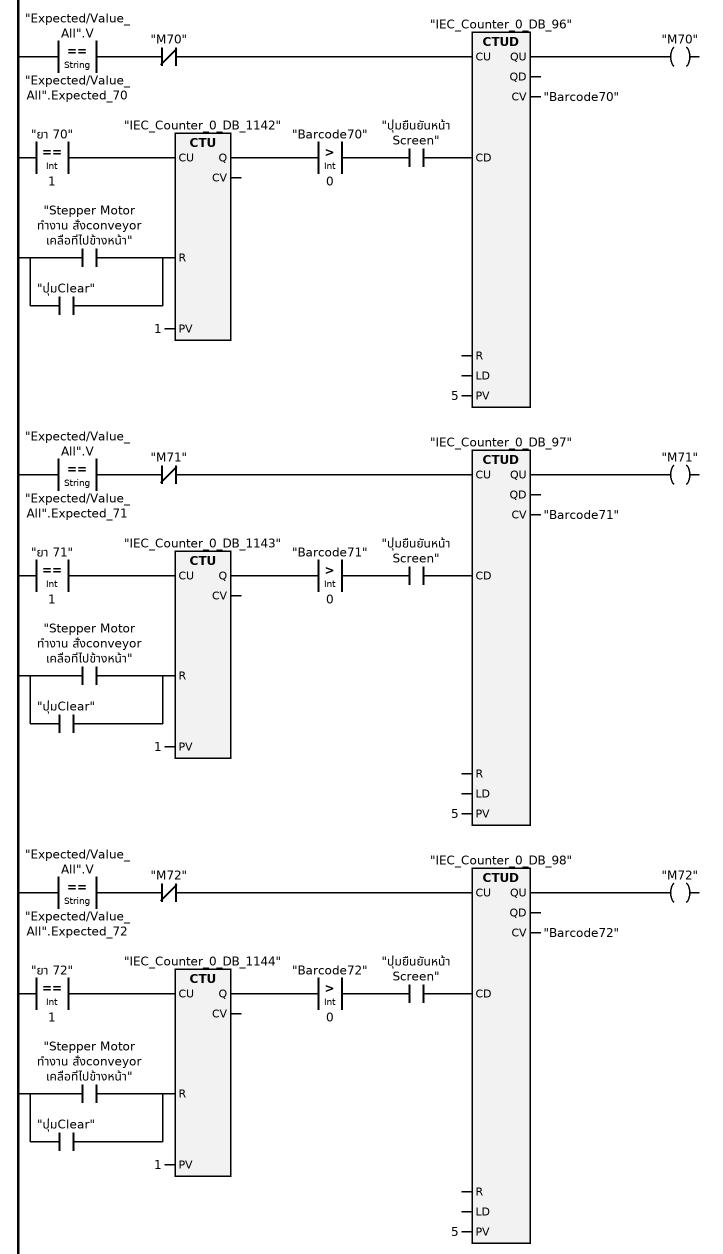
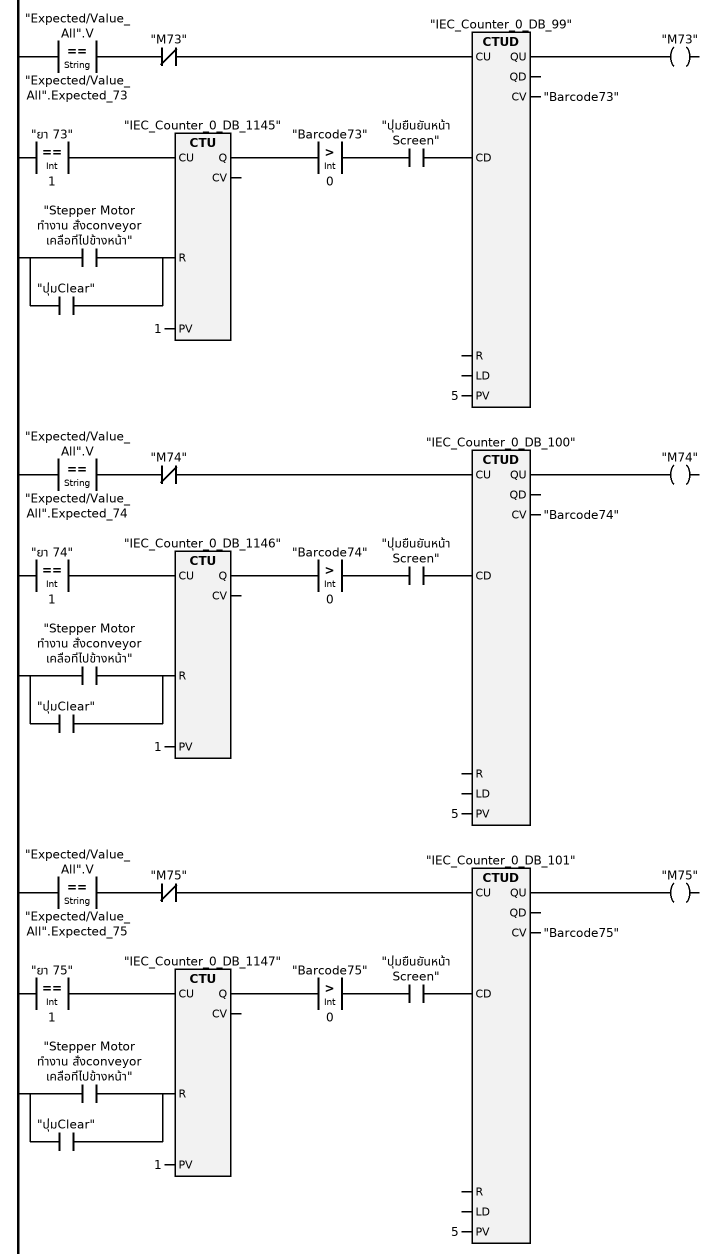
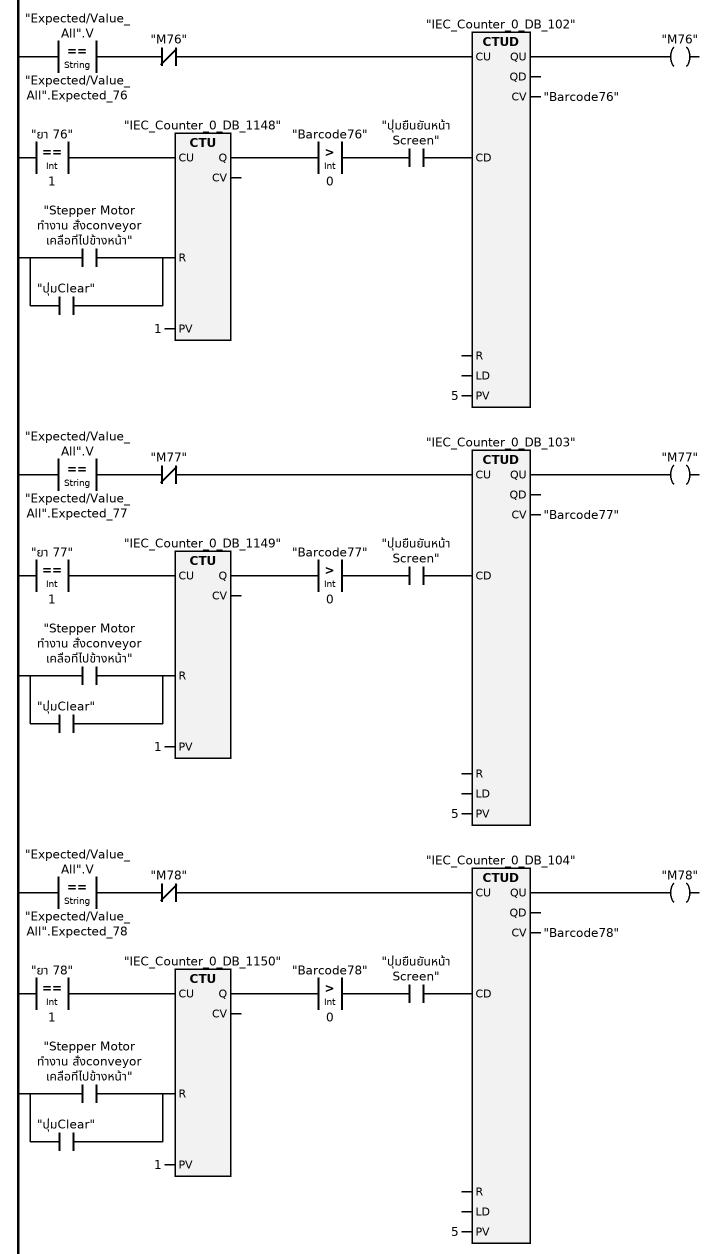
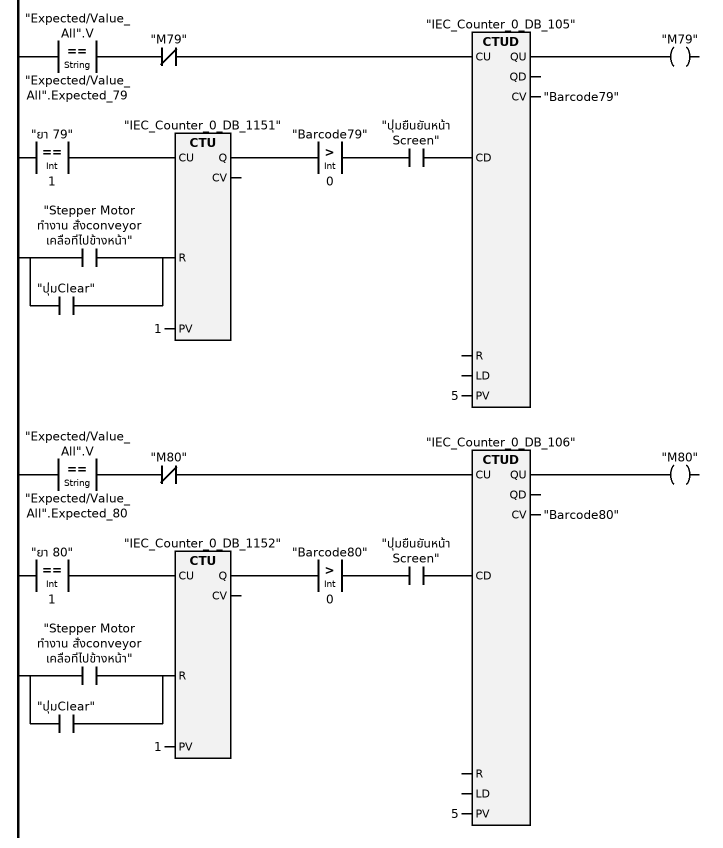
   "IEC_Counter_0_DB_1133".CTU(CU := "ยา 61" = 1,
                           R := "Stepper Motor ทำงาน สั่งconveyor เคลื่อที่ไปข้างหน้า" OR "ปุ่มClear",
                           PV := 1);
   "IEC_Counter_0_DB_87".CTUD(CU := ("Expected/Value_All".V = "Expected/Value_All".Expected_61) AND NOT "M61",
                           CD := "IEC_Counter_0_DB_1133".Q AND ("Barcode61" > 0) AND "ปุ่มยืนยันหน้า Screen",
                           PV := 5,
                           CV => "Barcode61");
   "M61" := "IEC_Counter_0_DB_87".QU;
   "IEC_Counter_0_DB_1134".CTU(CU := "ยา 62" = 1,
                           R := "Stepper Motor ทำงาน สั่งconveyor เคลื่อที่ไปข้างหน้า" OR "ปุ่มClear",
                           PV := 1);
   "IEC_Counter_0_DB_88".CTUD(CU := ("Expected/Value_All".V = "Expected/Value_All".Expected_62) AND NOT "M62",
                           CD := "IEC_Counter_0_DB_1134".Q AND ("Barcode62" > 0) AND "ปุ่มยืนยันหน้า Screen",
                           PV := 5,
                           CV => "Barcode62");
   "M62" := "IEC_Counter_0_DB_88".QU;
   "IEC_Counter_0_DB_1135".CTU(CU := "ยา 63" = 1,
                           R := "Stepper Motor ทำงาน สั่งconveyor เคลื่อที่ไปข้างหน้า" OR "ปุ่มClear",
                           PV := 1);
   "IEC_Counter_0_DB_89".CTUD(CU := ("Expected/Value_All".V = "Expected/Value_All".Expected_63) AND NOT "M63",
                           CD := "IEC_Counter_0_DB_1135".Q AND ("Barcode63" > 0) AND "ปุ่มยืนยันหน้า Screen",
                           PV := 5,
                           CV => "Barcode63");
   "M63" := "IEC_Counter_0_DB_89".QU;
   "IEC_Counter_0_DB_1136".CTU(CU := "ยา 64" = 1,
                           R := "Stepper Motor ทำงาน สั่งconveyor เคลื่อที่ไปข้างหน้า" OR "ปุ่มClear",
                           PV := 1);
   "IEC_Counter_0_DB_90".CTUD(CU := ("Expected/Value_All".V = "Expected/Value_All".Expected_64) AND NOT "M64",
                           CD := "IEC_Counter_0_DB_1136".Q AND ("Barcode64" > 0) AND "ปุ่มยืนยันหน้า Screen",
                           PV := 5,
                           CV => "Barcode64");
   "M64" := "IEC_Counter_0_DB_90".QU;
   "IEC_Counter_0_DB_1137".CTU(CU := "ยา 65" = 1,
                           R := "Stepper Motor ทำงาน สั่งconveyor เคลื่อที่ไปข้างหน้า" OR "ปุ่มClear",
                           PV := 1);
   "IEC_Counter_0_DB_91".CTUD(CU := ("Expected/Value_All".V = "Expected/Value_All".Expected_65) AND NOT "M65",
                           CD := "IEC_Counter_0_DB_1137".Q AND ("Barcode65" > 0) AND "ปุ่มยืนยันหน้า Screen",
                           PV := 5,
                           CV => "Barcode65");
   "M65" := "IEC_Counter_0_DB_91".QU;
   "IEC_Counter_0_DB_1138".CTU(CU := "ยา 66" = 1,
                           R := "Stepper Motor ทำงาน สั่งconveyor เคลื่อที่ไปข้างหน้า" OR "ปุ่มClear",
                           PV := 1);
   "IEC_Counter_0_DB_92".CTUD(CU := ("Expected/Value_All".V = "Expected/Value_All".Expected_66) AND NOT "M66",
                           CD := "IEC_Counter_0_DB_1138".Q AND ("Barcode66" > 0) AND "ปุ่มยืนยันหน้า Screen",
                           PV := 5,
                           CV => "Barcode66");
   "M66" := "IEC_Counter_0_DB_92".QU;
   "IEC_Counter_0_DB_1139".CTU(CU := "ยา 67" = 1,
                           R := "Stepper Motor ทำงาน สั่งconveyor เคลื่อที่ไปข้างหน้า" OR "ปุ่มClear",
                           PV := 1);
   "IEC_Counter_0_DB_93".CTUD(CU := ("Expected/Value_All".V = "Expected/Value_All".Expected_67) AND NOT "M67",
                           CD := "IEC_Counter_0_DB_1139".Q AND ("Barcode67" > 0) AND "ปุ่มยืนยันหน้า Screen",
                           PV := 5,
                           CV => "Barcode67");
   "M67" := "IEC_Counter_0_DB_93".QU;
   "IEC_Counter_0_DB_1140".CTU(CU := "ยา 68" = 1,
                           R := "Stepper Motor ทำงาน สั่งconveyor เคลื่อที่ไปข้างหน้า" OR "ปุ่มClear",
                           PV := 1);
   "IEC_Counter_0_DB_94".CTUD(CU := ("Expected/Value_All".V = "Expected/Value_All".Expected_68) AND NOT "M68",
                           CD := "IEC_Counter_0_DB_1140".Q AND ("Barcode68" > 0) AND "ปุ่มยืนยันหน้า Screen",
                           PV := 5,
                           CV => "Barcode68");
   "M68" := "IEC_Counter_0_DB_94".QU;
   "IEC_Counter_0_DB_1141".CTU(CU := "ยา 69" = 1,
                           R := "Stepper Motor ทำงาน สั่งconveyor เคลื่อที่ไปข้างหน้า" OR "ปุ่มClear",
                           PV := 1);
   "IEC_Counter_0_DB_95".CTUD(CU := ("Expected/Value_All".V = "Expected/Value_All".Expected_69) AND NOT "M69",
                           CD := "IEC_Counter_0_DB_1141".Q AND ("Barcode69" > 0) AND "ปุ่มยืนยันหน้า Screen",
                           PV := 5,
                           CV => "Barcode69");
   "M69" := "IEC_Counter_0_DB_95".QU;
   "IEC_Counter_0_DB_1142".CTU(CU := "ยา 70" = 1,
                           R := "Stepper Motor ทำงาน สั่งconveyor เคลื่อที่ไปข้างหน้า" OR "ปุ่มClear",
                           PV := 1);
   "IEC_Counter_0_DB_96".CTUD(CU := ("Expected/Value_All".V = "Expected/Value_All".Expected_70) AND NOT "M70",
                           CD := "IEC_Counter_0_DB_1142".Q AND ("Barcode70" > 0) AND "ปุ่มยืนยันหน้า Screen",
                           PV := 5,
                           CV => "Barcode70");
   "M70" := "IEC_Counter_0_DB_96".QU;
   "IEC_Counter_0_DB_1143".CTU(CU := "ยา 71" = 1,
                           R := "Stepper Motor ทำงาน สั่งconveyor เคลื่อที่ไปข้างหน้า" OR "ปุ่มClear",
                           PV := 1);
   "IEC_Counter_0_DB_97".CTUD(CU := ("Expected/Value_All".V = "Expected/Value_All".Expected_71) AND NOT "M71",
                           CD := "IEC_Counter_0_DB_1143".Q AND ("Barcode71" > 0) AND "ปุ่มยืนยันหน้า Screen",
                           PV := 5,
                           CV => "Barcode71");
   "M71" := "IEC_Counter_0_DB_97".QU;
   "IEC_Counter_0_DB_1144".CTU(CU := "ยา 72" = 1,
                           R := "Stepper Motor ทำงาน สั่งconveyor เคลื่อที่ไปข้างหน้า" OR "ปุ่มClear",
                           PV := 1);
   "IEC_Counter_0_DB_98".CTUD(CU := ("Expected/Value_All".V = "Expected/Value_All".Expected_72) AND NOT "M72",
                           CD := "IEC_Counter_0_DB_1144".Q AND ("Barcode72" > 0) AND "ปุ่มยืนยันหน้า Screen",
                           PV := 5,
                           CV => "Barcode72");
   "M72" := "IEC_Counter_0_DB_98".QU;
   "IEC_Counter_0_DB_1145".CTU(CU := "ยา 73" = 1,
                           R := "Stepper Motor ทำงาน สั่งconveyor เคลื่อที่ไปข้างหน้า" OR "ปุ่มClear",
                           PV := 1);
   "IEC_Counter_0_DB_99".CTUD(CU := ("Expected/Value_All".V = "Expected/Value_All".Expected_73) AND NOT "M73",
                           CD := "IEC_Counter_0_DB_1145".Q AND ("Barcode73" > 0) AND "ปุ่มยืนยันหน้า Screen",
                           PV := 5,
                           CV => "Barcode73");
   "M73" := "IEC_Counter_0_DB_99".QU;
   "IEC_Counter_0_DB_1146".CTU(CU := "ยา 74" = 1,
                           R := "Stepper Motor ทำงาน สั่งconveyor เคลื่อที่ไปข้างหน้า" OR "ปุ่มClear",
                           PV := 1);
   "IEC_Counter_0_DB_100".CTUD(CU := ("Expected/Value_All".V = "Expected/Value_All".Expected_74) AND NOT "M74",
                           CD := "IEC_Counter_0_DB_1146".Q AND ("Barcode74" > 0) AND "ปุ่มยืนยันหน้า Screen",
                           PV := 5,
                           CV => "Barcode74");
   "M74" := "IEC_Counter_0_DB_100".QU;
   "IEC_Counter_0_DB_1147".CTU(CU := "ยา 75" = 1,
                           R := "Stepper Motor ทำงาน สั่งconveyor เคลื่อที่ไปข้างหน้า" OR "ปุ่มClear",
                           PV := 1);
   "IEC_Counter_0_DB_101".CTUD(CU := ("Expected/Value_All".V = "Expected/Value_All".Expected_75) AND NOT "M75",
                           CD := "IEC_Counter_0_DB_1147".Q AND ("Barcode75" > 0) AND "ปุ่มยืนยันหน้า Screen",
                           PV := 5,
                           CV => "Barcode75");
   "M75" := "IEC_Counter_0_DB_101".QU;
   "IEC_Counter_0_DB_1148".CTU(CU := "ยา 76" = 1,
                           R := "Stepper Motor ทำงาน สั่งconveyor เคลื่อที่ไปข้างหน้า" OR "ปุ่มClear",
                           PV := 1);
   "IEC_Counter_0_DB_102".CTUD(CU := ("Expected/Value_All".V = "Expected/Value_All".Expected_76) AND NOT "M76",
                           CD := "IEC_Counter_0_DB_1148".Q AND ("Barcode76" > 0) AND "ปุ่มยืนยันหน้า Screen",
                           PV := 5,
                           CV => "Barcode76");
   "M76" := "IEC_Counter_0_DB_102".QU;
   "IEC_Counter_0_DB_1149".CTU(CU := "ยา 77" = 1,
                           R := "Stepper Motor ทำงาน สั่งconveyor เคลื่อที่ไปข้างหน้า" OR "ปุ่มClear",
                           PV := 1);
   "IEC_Counter_0_DB_103".CTUD(CU := ("Expected/Value_All".V = "Expected/Value_All".Expected_77) AND NOT "M77",
                           CD := "IEC_Counter_0_DB_1149".Q AND ("Barcode77" > 0) AND "ปุ่มยืนยันหน้า Screen",
                           PV := 5,
                           CV => "Barcode77");
   "M77" := "IEC_Counter_0_DB_103".QU;
   "IEC_Counter_0_DB_1150".CTU(CU := "ยา 78" = 1,
                           R := "Stepper Motor ทำงาน สั่งconveyor เคลื่อที่ไปข้างหน้า" OR "ปุ่มClear",
                           PV := 1);
   "IEC_Counter_0_DB_104".CTUD(CU := ("Expected/Value_All".V = "Expected/Value_All".Expected_78) AND NOT "M78",
                           CD := "IEC_Counter_0_DB_1150".Q AND ("Barcode78" > 0) AND "ปุ่มยืนยันหน้า Screen",
                           PV := 5,
                           CV => "Barcode78");
   "M78" := "IEC_Counter_0_DB_104".QU;
   "IEC_Counter_0_DB_1151".CTU(CU := "ยา 79" = 1,
                           R := "Stepper Motor ทำงาน สั่งconveyor เคลื่อที่ไปข้างหน้า" OR "ปุ่มClear",
                           PV := 1);
   "IEC_Counter_0_DB_105".CTUD(CU := ("Expected/Value_All".V = "Expected/Value_All".Expected_79) AND NOT "M79",
                           CD := "IEC_Counter_0_DB_1151".Q AND ("Barcode79" > 0) AND "ปุ่มยืนยันหน้า Screen",
                           PV := 5,
                           CV => "Barcode79");
   "M79" := "IEC_Counter_0_DB_105".QU;
   "IEC_Counter_0_DB_1152".CTU(CU := "ยา 80" = 1,
                           R := "Stepper Motor ทำงาน สั่งconveyor เคลื่อที่ไปข้างหน้า" OR "ปุ่มClear",
                           PV := 1);
   "IEC_Counter_0_DB_106".CTUD(CU := ("Expected/Value_All".V = "Expected/Value_All".Expected_80) AND NOT "M80",
                           CD := "IEC_Counter_0_DB_1152".Q AND ("Barcode80" > 0) AND "ปุ่มยืนยันหน้า Screen",
                           PV := 5,
                           CV => "Barcode80");
   "M80" := "IEC_Counter_0_DB_106".QU;
END_REGION

REGION Network 5
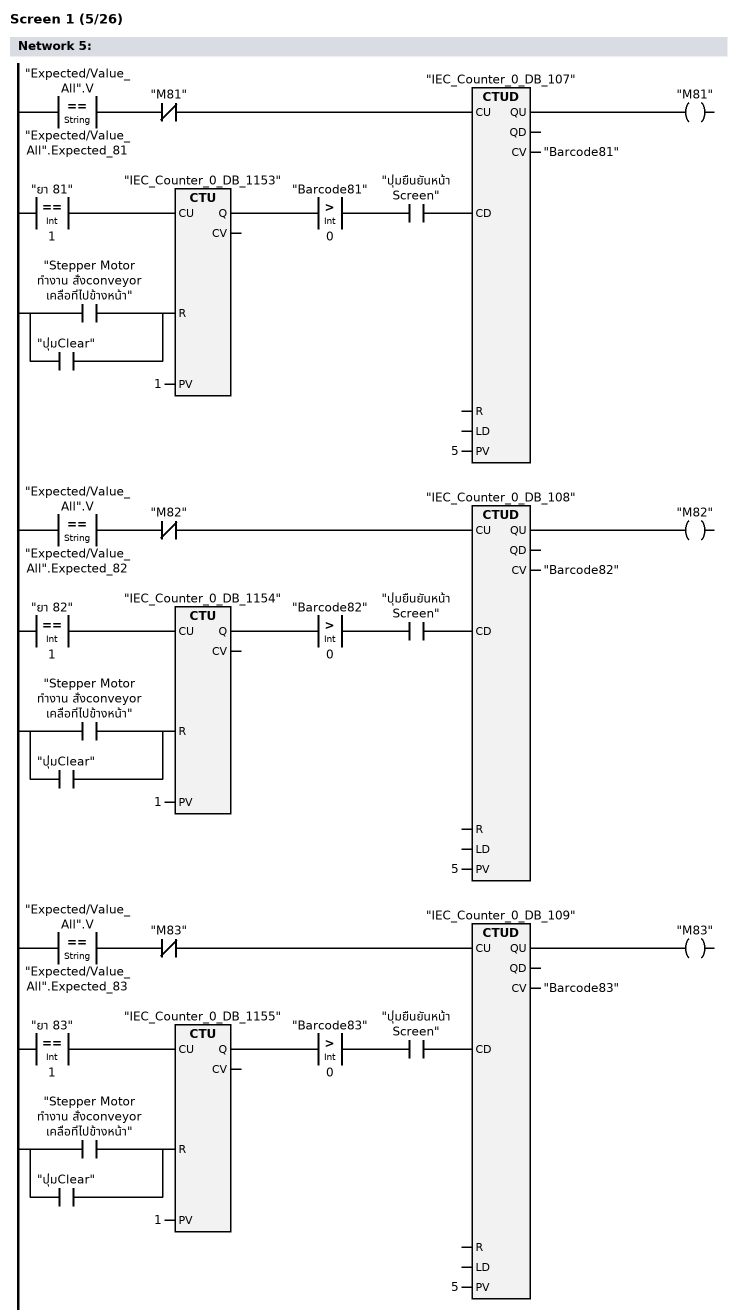
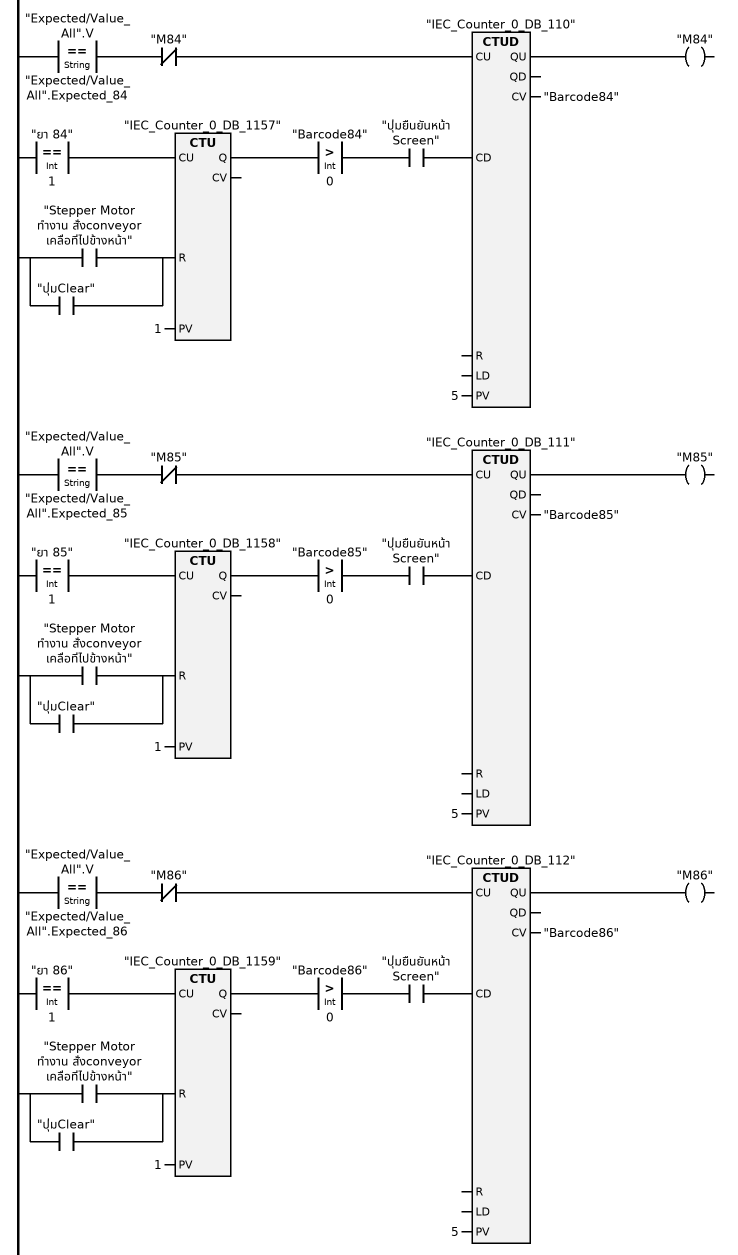
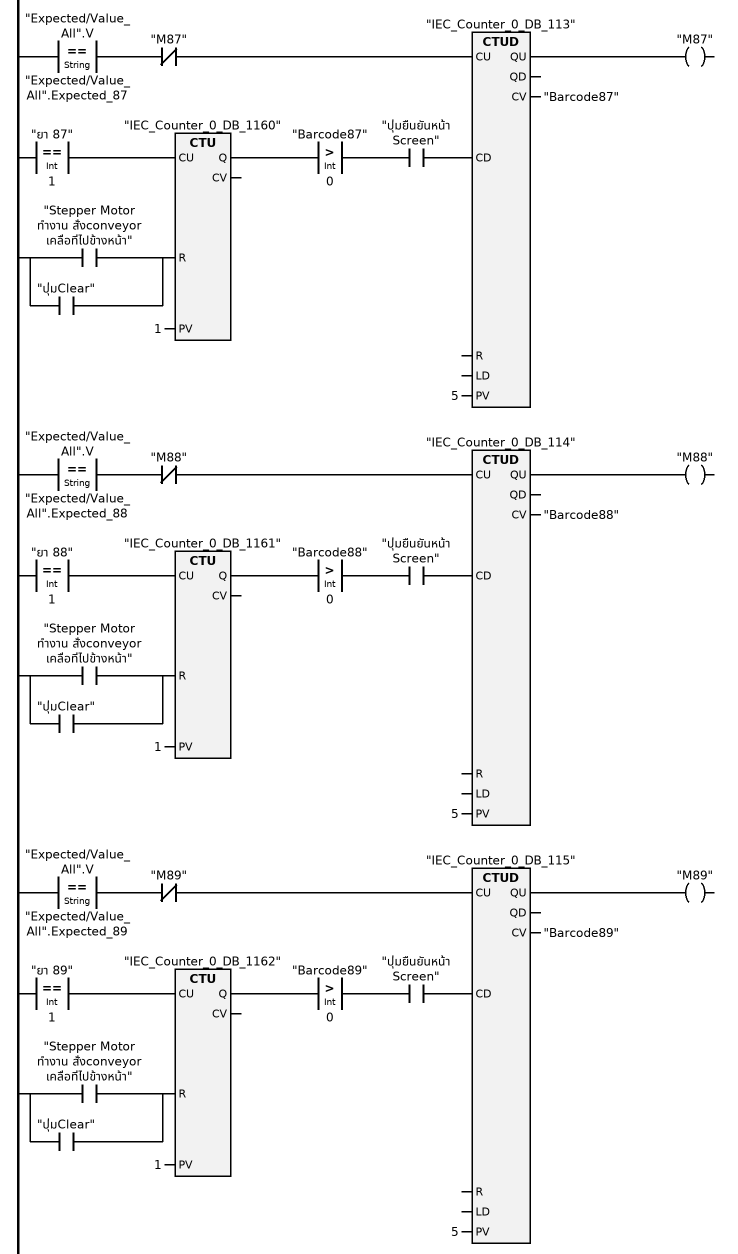
